// TwinCAT 3 PLC project PLC
// ProgramVersion: 3.1.4026.27
// libraries:
//   Tc2_Standard, * (Beckhoff Automation GmbH)
//   Tc2_System, * (Beckhoff Automation GmbH)
// project tree:
//   DUTs/ ST_EVENT.TcDUT
//   / PlcTask.TcTTO
//   POUs/FBs/ FB_SimEncoder.TcPOU
//   POUs/Function/ Celsius_To_Farenheit.TcPOU, Greater_Smaller.TcPOU, SwapNums.TcPOU
//   POUs/ MAIN.TcPOU, POU.TcPOU, TC3_Examples.TcPOU
// real-time tasks:
//   TASK PlcTask: cycle T#10ms, priority 6, ADS port 350

CONFIGURATION PLC
    RESOURCE PLC ON TwinCAT3
        TASK PlcTask(INTERVAL := T#10ms, PRIORITY := 6);
        PROGRAM MAIN WITH PlcTask : MAIN;
    END_RESOURCE
END_CONFIGURATION

// ---- DUTs/ST_EVENT.TcDUT
TYPE ST_EVENT : 
STRUCT
	eEventType : Tc2_System.TcEvent;
	eEventSeverity : Global.TcEventSeverity;
	nEventIdentity : UDINT;
	sEventText : STRING(255);
	dtTimeStamp : DATE_AND_TIME;
END_STRUCT
END_TYPE

// ---- POUs/MAIN.TcPOU
PROGRAM MAIN
VAR
    fbEnc : FB_SimEncoder;
    bGo   : BOOL;  // Wire to a HMI button or PLC tag
END_VAR

fbEnc(
    bActivate := bGo,
    rSpeed    := 1000.0,   // 1000 counts/s
    bDirection:= TRUE,
    nResolution := 4096    // e.g. 4096 PPR encoder
);

END_PROGRAM

// ---- POUs/FBs/FB_SimEncoder.TcPOU
FUNCTION_BLOCK FB_SimEncoder
VAR_INPUT
    bActivate   : BOOL;       // Set TRUE to start counting
    rSpeed      : LREAL := 0; // Encoder counts per second
    bDirection  : BOOL := TRUE; // TRUE = +, FALSE = -
    nResolution : UDINT := 4096; // Encoder PPR (for rollover)
END_VAR

VAR_OUTPUT
    nCount      : UDINT;      // Simulated encoder count (wraps at resolution)
    rPosition   : LREAL;      // Unwrapped position (in counts, signed)
    bRunning    : BOOL;       // TRUE while counting
END_VAR

VAR
    rDelta      : LREAL;      // Counts added this cycle
    rAccum      : LREAL := 0; // Accumulated (unwrapped) position
END_VAR

IF bActivate THEN
    bRunning := TRUE;

    // Calculate delta for this cycle (counts/s × cycle time)
	rDelta := rSpeed * (UDINT_TO_LREAL(_TaskInfo[GETCURTASKINDEXEX()].CycleTime) / 10_000_000.0);


    IF bDirection THEN
        rAccum := rAccum + rDelta;
    ELSE
        rAccum := rAccum - rDelta;
    END_IF

    // Wrap the UDINT count at the encoder resolution
	nCount := LREAL_TO_UDINT(rAccum) MOD nResolution;   

    // Unwrapped signed position
    rPosition := rAccum;

ELSE
    bRunning := FALSE;
    // Hold last values (no reset) — uncomment to reset:
    // nCount  := 0;
    // rPosition := 0;
    // rAccum  := 0;
END_IF

END_FUNCTION_BLOCK

// ---- POUs/Function/Celsius_To_Farenheit.TcPOU
FUNCTION Celsius_To_Farenheit : REAL
VAR_INPUT
	fCelsius : REAL;
END_VAR
VAR
END_VAR

Celsius_To_Farenheit := fCelsius * 1.8 + 32;

END_FUNCTION

// ---- POUs/Function/Greater_Smaller.TcPOU
FUNCTION Greater_Smaller : INT
VAR_INPUT
	nNumber1 : INT;
	nNumber2 : INT;
END_VAR
VAR_OUTPUT
	nGreater : INT;
	nSmaller : INT;
END_VAR

IF nNumber1 > nNumber2 THEN
	nGreater := nNumber1;
	nSmaller := nNumber2;
ELSE
	nGreater := nNumber2;
	nSmaller := nNumber1;
END_IF

END_FUNCTION

// ---- POUs/Function/SwapNums.TcPOU
FUNCTION SwapNums : INT
VAR_IN_OUT
	nNumber1 : INT;
	nNumber2 : INT;
END_VAR
VAR
	nNumberTemp : INT;
END_VAR

nNumberTemp := nNumber1;
nNumber1 := nNumber2;
nNumber2 := nNumberTemp;

END_FUNCTION

// ---- POUs/POU.TcPOU
PROGRAM POU
VAR
	fOneFloat : REAL;
	sThisIsAString : STRING;
	nAnInteger : INT;
	
	nReturnedNumberOfBytesForFloat : UDINT;
	nReturnedNumberOfBytesForString : UDINT;
	nReturnedNumberOfBytesForInteger : UDINT;
END_VAR

nReturnedNumberOfBytesForFloat := SIZEOF(fOneFloat);
nReturnedNumberOfBytesForString := SIZEOF(sThisIsAString);
nReturnedNumberOfBytesForInteger := SIZEOF(nAnInteger);

END_PROGRAM

// ---- POUs/TC3_Examples.TcPOU
PROGRAM TC3_Examples
VAR
	bOnlyRunOnce : BOOL;
	
	// Variables used to show how functions can operate
	fFarenheit : REAL;
	
	nReturnGreater : INT;
	nReturnSmaller : INT;
	
	nNumA : INT;
	nNumB : INT;
	
END_VAR

IF NOT bOnlyRunOnce THEN
	Tc2_System.ADSLOGSTR(msgCtrlMask := Tc2_System.Global_Variables.ADSLOG_MSGTYPE_ERROR OR Tc2_System.Global_Variables.ADSLOG_MSGTYPE_LOG,
						msgFmtStr := 'Hello World!',
						strArg := '');
	bOnlyRunOnce := TRUE;
END_IF

fFarenheit := Celsius_To_Farenheit(fCelsius := 5.0);

Greater_Smaller(nNumber1 := 2, nNumber2 := 9, nGreater => nReturnGreater, nSmaller => nReturnSmaller);

SwapNums(nNumA, nNumB);

POU();

END_PROGRAM
